// TIA Portal V19 export
DATA_BLOCK "RecipeActive"   // DB26
{ S7_Optimized_Access := 'TRUE' }
// stored: MemoryReserve 100
   VAR
      PositionsOffsetRobot_1 : Array[0..7] of "ST_TPM_AutoPosition";
   END_VAR
BEGIN
END_DATA_BLOCK
